Fanuc KAREL source: kx00005.KL

PROGRAM KX00005
%STACKSIZE=65535
%PRIORITY=65535
%NOLOCKGROUP
VAR
I : INTEGER
J : INTEGER
B : BOOLEAN
F : FILE
S : STRING[80]
P : XYZWPR
BEGIN
OPEN FILE F ('RW','MD:KFSAMPLE.DT')
-- UNRESOLVED_PC line 12 opcodes [22 A3] marker_code=32
CLOSE FILE F
END KX00005
